(* IEC 61131-3 sources: llm-plc-st-eval/data/processed_definitivo/gemini-3.1-pro-preview/B6/few_shot, 3 files *)

(* ---- ejec_1.st ---- *)
FUNCTION_BLOCK FB_Baliza
VAR_INPUT
    alarma : BOOL; (* Condicion de alarma *)
END_VAR
VAR_OUTPUT
    lampara : BOOL; (* Lampara de la baliza *)
END_VAR
VAR
    tOn : TON; (* Temporizador de fase encendida *)
    tOff : TON; (* Temporizador de fase apagada *)
END_VAR

(* Generador de intermitencia: 1s ON y 1s OFF mientras la alarma este activa *)
tOn(IN := alarma AND NOT tOff.Q, PT := T#1S);
tOff(IN := tOn.Q, PT := T#1S);

(* La lampara se enciende inmediatamente con la alarma y alterna su estado *)
lampara := alarma AND NOT tOn.Q;
END_FUNCTION_BLOCK

(* ---- ejec_2.st ---- *)
FUNCTION_BLOCK FB_Baliza
VAR_INPUT
    alarma : BOOL; (* Condicion de alarma *)
END_VAR
VAR_OUTPUT
    lampara : BOOL; (* Lampara de la baliza *)
END_VAR
VAR
    tonOn : TON; (* Temporizador de fase encendida *)
    tonOff : TON; (* Temporizador de fase apagada *)
END_VAR

(* Generador de pulsos: alterna entre temporizadores cada 1 segundo *)
tonOn(IN := alarma AND NOT tonOff.Q, PT := T#1S);
tonOff(IN := tonOn.Q, PT := T#1S);

(* La lampara enciende inmediatamente con la alarma y parpadea 1s ON / 1s OFF *)
lampara := alarma AND NOT tonOn.Q;
END_FUNCTION_BLOCK

(* ---- ejec_3.st ---- *)
FUNCTION_BLOCK FB_Baliza
VAR_INPUT
    alarma : BOOL; (* Condicion de alarma *)
END_VAR
VAR_OUTPUT
    lampara : BOOL; (* Lampara de la baliza *)
END_VAR
VAR
    tEncendido : TON; (* Temporizador de fase encendida *)
    tApagado : TON; (* Temporizador de fase apagada *)
END_VAR

(* Ciclo de parpadeo: 1s encendido, 1s apagado mientras la alarma este activa *)
tEncendido(IN := alarma AND NOT tApagado.Q, PT := T#1S);
tApagado(IN := tEncendido.Q, PT := T#1S);

(* La lampara enciende inmediatamente con la alarma y alterna su estado cada segundo *)
lampara := alarma AND NOT tEncendido.Q;
END_FUNCTION_BLOCK
